// TIA Portal V20 export
ORGANIZATION_BLOCK "T12_Ciclo"   // OB132, LAD, ProgramCycle
TITLE = T12_Ciclo
{ S7_Optimized_Access := 'TRUE' }
AUTHOR : IA
FAMILY : PRUEBA
VERSION : 0.1
// Tanda 7: llama a las pruebas
// stored: AutoNumber false, IsIECCheckEnabled false, SetENOAutomatically false
   VAR_INPUT
      Initial_Call : Bool;
      Remanence : Bool;
   END_VAR
BEGIN

REGION Network 1: T12_S_Pruebas
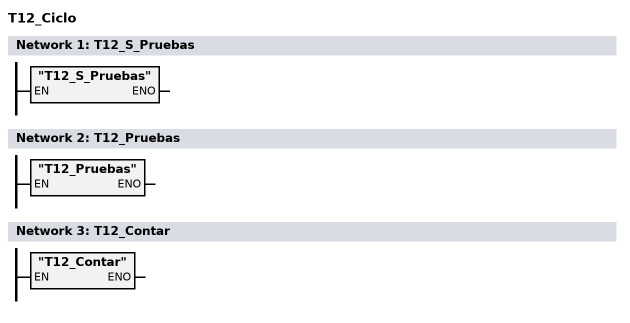
   RUNG wire#powerrail
      "T12_S_Pruebas"()
   END_RUNG
   // the same network as SCL:
   "T12_S_Pruebas"();
END_REGION

REGION Network 2: T12_Pruebas
   RUNG wire#powerrail
      "T12_Pruebas"()
   END_RUNG
   // the same network as SCL:
   "T12_Pruebas"();
END_REGION

REGION Network 3: T12_Contar
   RUNG wire#powerrail
      "T12_Contar"()
   END_RUNG
   // the same network as SCL:
   "T12_Contar"();
END_REGION
END_ORGANIZATION_BLOCK
